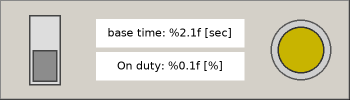
VISUALIZATION vis_FB_DutyCycle  // 350x100
VAR_IN_OUT
	fb: FB_DutyCycle;
END_VAR
    Rectangle (0,0 350x100)
    Lamp1 (266,15 70x70), variable: fb.bOut, style: Lamp-Lamp1-Yellow
    DipSwitch (10,15 70x70), variable: fb.bEnable, behaviour: TOGGLE, style: Switch-DipSwitch-Gray
    Textfield (95,18 150x30), "base time: %2.1f [sec]", text variable: fb.fBaseTime, input disabled if: prg_User.actUser<4
        OnMouseClick: write the text variable via Edit, min 0, max 60
    Textfield (95,51 150x30), "On duty: %0.1f [%]", text variable: fb.fOn_Duty
        OnMouseClick: write the text variable via Edit, min 0, max 100
END_VISUALIZATION

(* stored: Version 1.1.0.1, ProductVersion 3.1.4024.12
   Visu vis_FB_DutyCycle: Id {8c91fbb2-1ca9-4bed-85da-f49f29b5cfd6} *)
